TYPE "naut_Motor"
VERSION : 0.1
   STRUCT
      Run : BOOL;
      Speed : REAL;
   END_STRUCT;

END_TYPE
